TYPE ST_PeelerToUnity :
STRUCT
	fY          : REAL;    // Y position (0 - 100%)
	GameIsActive : BOOL;
   

END_STRUCT
END_TYPE

(* stored: Version 1.1.0.1, ProductVersion 3.1.4024.15
   DUT ST_PeelerToUnity: Id {fe2805ba-2128-4d98-b4ac-0aff45629c3c} *)
